Fanuc KAREL source: kd00013.KL

-- PROVISIONAL review KL for V1013-1; original PC SHA256 3ba56fb99c9466fd0ee1aa6cedf932686824814c7e4a810ff2186c621333c65f
-- Incomplete behavior may be omitted. Consult companion uncertainty JSON. Do not deploy.
PROGRAM KD00013
%NOLOCKGROUP
VAR
  I : INTEGER
  J : INTEGER
  B : BOOLEAN
  R : REAL
  S : STRING[80]
BEGIN
  -- UNRESOLVED_PC offsets 5-13; opcodes 2E,9D,1A
  -- UNRESOLVED_PC offsets 18-22; opcodes 7F
END KD00013
